Staubli VAL3: Lab2A_L2.pjx

--- Lab2A_L2.pjx ---
parameters version=s6.8 stackSize=5000 millimeterUnit=true
program file=start.pgx
program file=pickAndPlace.pgx
program file=stop.pgx
program file=physicalIO.pgx
data file=Lab2A_L2.dtx
alias name=io interface=io autoload=true

--- Lab2A_L2.dtx ---


--- start.pgx ---
program start()
// Lab2A Level 2 - parts loaded in ramps
  local num rowIndex
  local num columnIndex
  local num targetIndex
  local pointRs targetPose
begin
  // Four parts in each ramp. Start with an empty matrix.
  userPage()
  cls()
  physicalRun = !simulation
  cycleStep = 0
  vacuumOn = false
  blowOn = false
  ioReady = false

  if physicalRun
    taskCreate "physicalIO", 10, physicalIO()
    wait(ioReady == true)
    putln("PHYSICAL - parts loaded in ramps")
  else
    putln("SIMULATION - edit partOnTool at steps 60 and 70")
  endIf

  moveSpeed.vel = 10
  moveSpeed.accel = 10
  moveSpeed.decel = 10
  moveSpeed.blend = off

  // Each row starts at its own taught pose (0 or 4).
  for rowIndex = 0 to 1
    for columnIndex = 0 to 3
      targetIndex = 4*rowIndex + columnIndex
      targetPose = jointToPoint(vacuumTool, world, placePose[4*rowIndex])
      targetPose.trsf.y = targetPose.trsf.y + 60*columnIndex
      if columnIndex != 0
        if !pointToJoint(vacuumTool, placePose[4*rowIndex], targetPose, placePose[targetIndex])
          putln("ERROR: unreachable matrix destination")
          putln(targetIndex)
          return
        endIf
      endIf

      targetPose.trsf.z = targetPose.trsf.z + 50
      if !pointToJoint(vacuumTool, placePose[targetIndex], targetPose, placeApproach[targetIndex])
        putln("ERROR: unreachable matrix approach")
        putln(targetIndex)
        return
      endIf
    endFor
  endFor

  movej(homePose, vacuumTool, moveSpeed)
  waitEndMove()

  // Alternate ramps for each column: 0,4,1,5,2,6,3,7.
  for columnIndex = 0 to 3
    for materialType = 0 to 1
      placeIndex = 4*materialType + columnIndex
      putln("Place in slot:")
      putln(placeIndex)
      call pickAndPlace()
    endFor
  endFor

  cycleStep = 100
  putln("Level 2 completed: eight parts placed")
end

--- physicalIO.pgx ---
program physicalIO()
// Suction tool inputs and outputs
begin
  // Only the suction tool is controlled in Levels 1 and 2.
  while true
    partOnTool = io:bIn0 == true
    io:bOut0 = vacuumOn
    io:bOut1 = blowOn
    ioReady = true
    delay(0.01)
  endWhile
end

--- pickAndPlace.pgx ---
program pickAndPlace()
// Pick one part, place it and return home
begin
  // materialType selects the ramp; placeIndex selects the destination.
  vacuumOn = false
  blowOn = false
  movej(pickApproach[materialType], vacuumTool, moveSpeed)
  waitEndMove()
  movel(jointToPoint(vacuumTool, world, pickPose[materialType]), vacuumTool, moveSpeed)
  waitEndMove()
  vacuumOn = true
  cycleStep = 60
  putln("60 - Wait for partOnTool=true")
  wait(partOnTool == true)
  movel(jointToPoint(vacuumTool, world, pickApproach[materialType]), vacuumTool, moveSpeed)
  waitEndMove()

  movej(placeApproach[placeIndex], vacuumTool, moveSpeed)
  waitEndMove()
  movel(jointToPoint(vacuumTool, world, placePose[placeIndex]), vacuumTool, moveSpeed)
  waitEndMove()
  vacuumOn = false
  blowOn = true
  delay(0.3)
  blowOn = false
  cycleStep = 70
  putln("70 - Wait for partOnTool=false")
  wait(partOnTool == false)

  movel(jointToPoint(vacuumTool, world, placeApproach[placeIndex]), vacuumTool, moveSpeed)
  waitEndMove()
  movej(homePose, vacuumTool, moveSpeed)
  waitEndMove()
end

--- stop.pgx ---
program stop()
// Stop motion and preserve suction
begin
  resetMotion()
  blowOn = false
  if physicalRun
    taskKill("physicalIO")
    io:bOut1 = false
  endIf
  // Preserve suction so a held part is not released by STOP.
  cycleStep = -1
  putln("Stopped - empty the destinations before restarting")
end
